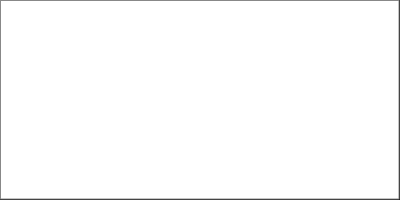
VISUALIZATION V_NCIMeina2_1000x1000_Circles  // 400x200
VAR_IN_OUT
	HMI : ST_PackMLBaseModule_HMI;
	HMI_GantryXYZ : ST_GantryXYZ_HMI;
	HMI_Recipe : ST_RecipeBuilder_HMI;
END_VAR
    RoundedRectangle (0,0 400x200)
END_VISUALIZATION

(* stored: Version 1.1.0.1, ProductVersion 3.1.4024.15
   Visu V_NCIMeina2_1000x1000_Circles: Id {ceb3d707-85b5-4ea5-bea9-aa2192732bf6} *)
